Fanuc KAREL source: kd00072.KL

-- PROVISIONAL review KL for V940-1; original PC SHA256 fa76f12ec1f2a71987c10a55701f14230f4de8badcda8a40dbb5c71f795dd76a
-- Incomplete behavior may be omitted. Consult companion uncertainty JSON. Do not deploy.
PROGRAM KD00072
%NOLOCKGROUP
VAR
  I : INTEGER
  J : INTEGER
  B : BOOLEAN
  R : REAL
  S : STRING[80]
BEGIN
  -- V9_IO_1F02_MOTIF_HINT bounded seven-record physical form; historical source, timing/runtime/producer release held
  -- V9_ZERO_TABLE_METADATA_HINT layout=0001; no indexed target words; source/name/runtime held
  -- UNRESOLVED_PC offsets 5-13; opcodes 9D,2E,1F
  -- UNRESOLVED_PC offsets 18-22; opcodes 7F
END KD00072
